TYPE ST_EL3356CoeWriteData_1 :
STRUCT
	wIdx: WORD;
	bySubIdx: BYTE;
	bWriteOK: BOOL;
	dwData: DWORD;
	nSize: UDINT;
END_STRUCT
END_TYPE

(* stored: Version 1.1.0.1, ProductVersion 3.1.4024.15
   DUT ST_EL3356CoeWriteData_1: Id {4ebf91c0-aded-41a8-a41c-8d732b5ddd39} *)
